// TIA Portal V20 export
// export: Created 2026-10-12T05:42:34.4093582Z, ExportSetting WithDefaults, DisplayName Totally Integrated Automation Portal, DisplayVersion V20, DisplayName TIA Portal Openness, DisplayVersion V20, DisplayName TIA Portal Teamcenter Gateway, DisplayVersion V20, DisplayName TIA Portal Version Control Interface, DisplayVersion V20, DisplayName SINAMICS Startdrive Advanced, DisplayVersion V20 SP1 Update 2, DisplayName SINAMICS Startdrive G110M, G120, G120C, G120D, G120P, G115D, DisplayVersion V20 SP1 Update 2, DisplayName SINAMICS Startdrive G130, G150, S120, S150, SINAMICS MV, G220, S200, S210, DisplayVersion V20 SP1 Update 2, DisplayName STEP 7 Professional, DisplayVersion V20, DisplayName STEP 7 Safety, DisplayVersion V20, DisplayName WinCC Basic/Comfort/Advanced, DisplayVersion V20, DisplayName WinCC Professional, DisplayVersion V20, DisplayName WinCC Unified, DisplayVersion V20
FUNCTION "F_PressDemoRamResult" : Void   // FC164, SCL
{ S7_Optimized_Access := 'TRUE' }
VERSION : 0.1
// stored: AutoNumber true, IsIECCheckEnabled false, SetENOAutomatically false, UDAEnableTagReadback false
   VAR_INPUT
      Reached : Bool;
   END_VAR
   VAR_IN_OUT
      Seq : "FRK_SequenceCtx";
      Cycle : "ST_PressDemoCycle";
      AlarmLog : "FRK_AlarmLog";
   END_VAR
BEGIN

   "FRK_SeqSelect"(Seq := #Seq,
                   AdvanceOk := #Reached,
                   Jump1Ok := #Seq.CommandFailed);
   IF #Seq.RetVal = 2 THEN
       #Cycle.FailureReason := #Seq.HandledDiagnostic.ReasonCode;
       "FRK_SeqMessage"(Seq := #Seq,
                        AlarmLog := #AlarmLog,
                        Diag := #Seq.HandledDiagnostic);
   END_IF;
END_FUNCTION
